(* IEC 61131-3 sources: llm-plc-st-eval/data/definitivo/claude-sonnet-4-6/B6/zero_shot, 3 files *)

(* ---- ejec_1.st ---- *)
```pascal
FUNCTION_BLOCK FB_Baliza
VAR_INPUT
    alarma : BOOL; (* Condición de alarma activa *)
END_VAR

VAR_OUTPUT
    lampara : BOOL; (* Salida de la lámpara de baliza *)
END_VAR

VAR
    tonEncendida : TON; (* Temporizador para tiempo encendida *)
    tonApagada   : TON; (* Temporizador para tiempo apagada *)
    estadoLuz    : BOOL; (* Estado interno del parpadeo: TRUE=encendida *)
END_VAR

(* ─────────────────────────────────────────────
   Lógica principal
   ───────────────────────────────────────────── *)

IF NOT alarma THEN
    (* Sin alarma: apagar lámpara y resetear todo *)
    lampara      := FALSE;
    estadoLuz    := FALSE;
    tonEncendida(IN := FALSE, PT := T#1S);
    tonApagada  (IN := FALSE, PT := T#1S);

ELSE
    (* Con alarma: alternar entre encendida y apagada *)

    IF estadoLuz THEN
        (* Fase encendida: esperar 1 s y luego pasar a apagada *)
        tonApagada  (IN := FALSE, PT := T#1S); (* Mantener apagado el otro TON *)
        tonEncendida(IN := TRUE,  PT := T#1S);

        IF tonEncendida.Q THEN
            (* Tiempo encendida cumplido → cambiar a fase apagada *)
            estadoLuz := FALSE;
            tonEncendida(IN := FALSE, PT := T#1S); (* Reset *)
        END_IF;

    ELSE
        (* Fase apagada: esperar 1 s y luego pasar a encendida *)
        tonEncendida(IN := FALSE, PT := T#1S); (* Mantener apagado el otro TON *)
        tonApagada  (IN := TRUE,  PT := T#1S);

        IF tonApagada.Q THEN
            (* Tiempo apagada cumplido → cambiar a fase encendida *)
            estadoLuz := TRUE;
            tonApagada(IN := FALSE, PT := T#1S); (* Reset *)
        END_IF;

    END_IF;

    (* La salida refleja el estado interno del parpadeo *)
    lampara := estadoLuz;

END_IF;
```

(* ---- ejec_2.st ---- *)
```pascal
FUNCTION_BLOCK FB_Baliza
VAR_INPUT
    alarma : BOOL; (* Condición de alarma activa *)
END_VAR

VAR_OUTPUT
    lampara : BOOL; (* Salida hacia la lámpara de baliza *)
END_VAR

VAR
    tonEncendido  : TON; (* Temporizador para tiempo encendida *)
    tonApagado    : TON; (* Temporizador para tiempo apagada *)
    estadoLampara : BOOL := FALSE; (* Estado interno del parpadeo *)
END_VAR

(* -------------------------------------------------------
   Lógica de baliza de alarma
   - Sin alarma : lámpara apagada, temporizadores reseteados
   - Con alarma : parpadeo 1s ON / 1s OFF
   ------------------------------------------------------- *)

IF NOT alarma THEN
    (* Sin alarma: apagar lámpara y resetear todo *)
    estadoLampara := FALSE;
    tonEncendido(IN := FALSE, PT := T#1S);
    tonApagado(IN := FALSE, PT := T#1S);

ELSE
    (* Con alarma: gestionar ciclo de parpadeo *)

    IF NOT estadoLampara THEN
        (* Fase APAGADA: esperar 1 segundo *)
        tonEncendido(IN := FALSE, PT := T#1S); (* Mantener reseteado *)
        tonApagado(IN := TRUE,  PT := T#1S);

        IF tonApagado.Q THEN
            (* Tiempo apagada cumplido: pasar a fase encendida *)
            estadoLampara := TRUE;
            tonApagado(IN := FALSE, PT := T#1S); (* Resetear temporizador *)
        END_IF;

    ELSE
        (* Fase ENCENDIDA: esperar 1 segundo *)
        tonApagado(IN := FALSE, PT := T#1S);  (* Mantener reseteado *)
        tonEncendido(IN := TRUE,  PT := T#1S);

        IF tonEncendido.Q THEN
            (* Tiempo encendida cumplido: pasar a fase apagada *)
            estadoLampara := FALSE;
            tonEncendido(IN := FALSE, PT := T#1S); (* Resetear temporizador *)
        END_IF;

    END_IF;

END_IF;

(* Asignar estado interno a la salida *)
lampara := estadoLampara;

END_FUNCTION_BLOCK
```

(* ---- ejec_3.st ---- *)
```pascal
FUNCTION_BLOCK FB_Baliza
VAR_INPUT
    alarma : BOOL; (* Condición de alarma activa *)
END_VAR

VAR_OUTPUT
    lampara : BOOL; (* Salida hacia la lámpara de baliza *)
END_VAR

VAR
    tonEncendido  : TON; (* Temporizador para tiempo encendida *)
    tonApagado    : TON; (* Temporizador para tiempo apagada *)
    estadoLampara : BOOL := FALSE; (* Estado interno del parpadeo *)
END_VAR

(* -------------------------------------------------------
   Lógica de baliza de alarma
   - Sin alarma: lámpara apagada, temporizadores reseteados
   - Con alarma:  parpadeo 1s ON / 1s OFF
   ------------------------------------------------------- *)

IF NOT alarma THEN
    (* Sin alarma: apagar lámpara y resetear todo *)
    estadoLampara := FALSE;
    tonEncendido(IN := FALSE, PT := T#1S);
    tonApagado(IN := FALSE, PT := T#1S);

ELSE
    (* Con alarma: máquina de estados de parpadeo *)

    IF NOT estadoLampara THEN
        (* Fase APAGADA: esperar 1 segundo *)
        tonEncendido(IN := FALSE, PT := T#1S); (* Mantener reseteado *)
        tonApagado(IN := TRUE,  PT := T#1S);

        IF tonApagado.Q THEN
            (* Tiempo apagada cumplido: pasar a fase encendida *)
            estadoLampara := TRUE;
            tonApagado(IN := FALSE, PT := T#1S); (* Resetear temporizador *)
        END_IF;

    ELSE
        (* Fase ENCENDIDA: esperar 1 segundo *)
        tonApagado(IN := FALSE, PT := T#1S);  (* Mantener reseteado *)
        tonEncendido(IN := TRUE,  PT := T#1S);

        IF tonEncendido.Q THEN
            (* Tiempo encendida cumplido: pasar a fase apagada *)
            estadoLampara := FALSE;
            tonEncendido(IN := FALSE, PT := T#1S); (* Resetear temporizador *)
        END_IF;

    END_IF;

END_IF;

(* Asignar estado interno a la salida *)
lampara := estadoLampara AND alarma;

END_FUNCTION_BLOCK
```
